(* IEC 61131-3 sources: SortJet_MasterSPS_Aufbau.fbsproj/08_POUs/Basis Funktionsbausteine, 5 files *)

(* ---- Ampel_FB.fb.st ---- *)
(* METADATA
{
	"v3Meta": {
		"objectGuid": "3b447e4d-6caa-4c98-ad2d-e4c3e81f2c59"
	}
}
*)
FUNCTION_BLOCK Ampel_FB
VAR_INPUT

  // BOOL
  bpAutomatikAktiv                : BOOL;
  bpSystemcheckAktiv              : BOOL;
  bpBetriebsstoppAktiv            : BOOL;
  bpInternerBetriebsstopp         : BOOL;
  bpHinweisFWEingriffErforderlich : BOOL;
  bpSignalExtern                  : BOOL; // Blau Dauerlicht (z. B. Faecherwagen bald voll); Eingriff erforderlich hat Vorrang (blinkt)

END_VAR
VAR_OUTPUT
END_VAR
VAR

  //BOOL
  blFlashbit    : BOOL;

  // BYTE
  bylShiftByte  : BYTE :=1;

  // WORD
  wlModus       : WORD;
  wlInitAmpel   : WORD;

  // INT
  ilIndex       : INT;

  // TRIGGER
  rtlInitAmpel  : R_TRIG;

  // BLINK
  Flasher       : BLINK;

END_VAR
VAR

  // HARDWARE AUSGAENGE
  out_bAmpelLeuchteRot     AT%Q* : BOOL;
  out_bAmpelLeuchteGelb    AT%Q* : BOOL;
  out_bAmpelLeuchteGruen   AT%Q* : BOOL;
  out_bAmpelLeuchteBlau    AT%Q* : BOOL;

END_VAR
//-------------------------------------------------------------------------------------------------
// BAUSTEIN: ANSTEUERUNG
//-------------------------------------------------------------------------------------------------
(* Hinweis:
   - Baustein zum Ansteuern der optischen Signale des Sortjet : AMPELN
*)
Flasher(ENABLE:= TRUE , TIMELOW:= t#0.2s, TIMEHIGH:= t#0.2s , OUT=> blFlashbit);
rtlInitAmpel(CLK:= blFlashbit );

out_bAmpelLeuchteBlau := SEL( bpHinweisFWEingriffErforderlich, bpSignalExtern, gbFlashbit02sec );

//  Zentral den OperatingMode bestimmen
IF ( NOT NotHalt.bpNotHaltOK) THEN // NotAus nicht OK
  wlModus := 3;
ELSIF ( bpBetriebsstoppAktiv  ) THEN // Betriebsstop gesetzt
  wlModus := 8;
ELSIF ( Visu_Start_Auto ) THEN // VisuAuto aktiv
  wlModus := 7;
ELSIF ( bgInbetriebnahmeBit ) THEN // Inbetriebnahmebit gesetzt
  wlModus := 5;
ELSIF ( bpInternerBetriebsstopp ) THEN // Fehler/interner betriebsstop gesetzt
  wlModus := 0;
ELSIF ( Initialisierung.bpInitialisierungAktiv ) THEN // Initialiesierung aktiv
  wlModus := 5;
ELSIF ( bpSystemcheckAktiv ) THEN // Checkroutine aktiv
  wlModus := 6;
ELSIF ( bpAutomatikAktiv ) THEN // automatik aktiv
  wlModus := 2;
ELSE // Handbetrieb aktiv
  wlModus := 4;
END_IF

CASE wlModus OF
  // ======================================================
  0 : // Faliure active
    out_bAmpelLeuchteRot    := blFlashbit;
    out_bAmpelLeuchteGelb   := NOT out_bAmpelLeuchteRot;
    out_bAmpelLeuchteGruen  := FALSE;

  // ======================================================
  1:  // Service Mode
    out_bAmpelLeuchteRot    := FALSE;
    out_bAmpelLeuchteGelb   := TRUE;
    out_bAmpelLeuchteGruen  := FALSE;

  // ======================================================
  2:  // Automatic Running
    out_bAmpelLeuchteRot    := FALSE;
    out_bAmpelLeuchteGelb   := FALSE;
    out_bAmpelLeuchteGruen  := TRUE;

  // ======================================================
  3:  // Emergency Stop Active
    out_bAmpelLeuchteRot    := TRUE;
    out_bAmpelLeuchteGelb   := FALSE;
    out_bAmpelLeuchteGruen  := FALSE;

  // ======================================================
  4:   // Manual Mode
    out_bAmpelLeuchteRot    := FALSE;
    out_bAmpelLeuchteGelb   := TRUE;
    out_bAmpelLeuchteGruen  := FALSE;

  // ======================================================
  5: // Initialisation Mode
    out_bAmpelLeuchteRot    := ((wlInitAmpel AND Maske_Bit_2)<>0);
    out_bAmpelLeuchteGelb   :=((wlInitAmpel AND Maske_Bit_1)<>0);
    out_bAmpelLeuchteGruen  :=((wlInitAmpel AND Maske_Bit_0)<>0);

  // ======================================================
  6:   // Check Routine wurde gestartet
    out_bAmpelLeuchteRot    := FALSE;
    out_bAmpelLeuchteGelb   := FALSE;
    out_bAmpelLeuchteGruen  := blFlashbit;

  // ======================================================
  7:   // VisuAuto aktiv
    out_bAmpelLeuchteRot    := FALSE;
    out_bAmpelLeuchteGelb   := NOT blFlashbit;
    out_bAmpelLeuchteGruen  := TRUE;
  // ======================================================
  8:   // Betriebsstoptaster betätigt
    out_bAmpelLeuchteRot    := FALSE;
    out_bAmpelLeuchteGelb   := blFlashbit;
    out_bAmpelLeuchteGruen  := bpAutomatikAktiv;

// ======================================================
END_CASE

IF ( wlModus = 5) THEN

  IF ( rtlInitAmpel.Q ) THEN

    wlInitAmpel :=SHL(bylShiftByte, ilIndex);
    ilIndex := ilIndex + 1;

    IF ( ilIndex = 3 ) THEN
      ilIndex := 0;
    END_IF;

  END_IF;

ELSE
  wlInitAmpel := 0;

END_IF
END_FUNCTION_BLOCK

(* ---- BetriebsStop_FB.fb.st ---- *)
(* METADATA
{
	"v3Meta": {
		"objectGuid": "07d57a24-f3c0-4742-8d44-44a8d21cf93a"
	}
}
*)
FUNCTION_BLOCK BetriebsStop_FB
VAR_INPUT
END_VAR
VAR_OUTPUT

  // BOOLEAN
  abpBetriebsstop  : ARRAY [cERSTER_AUTOMATIKKREIS..cLETZTER_AUTOMATIKKREIS] OF BOOL;

END_VAR
VAR

  // BOOLEAN
  blBetriebsstop  : BOOL; // Merkervariable

  // WORD
  wlIndex                    : WORD;
  wMeldungsNrInkrementieren  : WORD := 0;

END_VAR
//-------------------------------------------------------------------------------------------------
// BAUSTEIN: BETRIEBSSTATUS
//-------------------------------------------------------------------------------------------------

(* Hinweis:
   - Betriebs- Stopp ausloesen
   - Internen Betriebsstop ausloesen
*)

blBetriebsstop := (  ( NOT bgMMIOK AND NOT bgMMIBruecken ) );

//-------------------------------------------------------------------------------------------------
// BAUSTEIN: MELDUNGEN
//-------------------------------------------------------------------------------------------------
(* Hinweis:
   - Generieren einer Meldung
*)
wMeldungsNrInkrementieren := 0;

FOR wlIndex := cERSTER_AUTOMATIKKREIS TO cLETZTER_AUTOMATIKKREIS DO
  abpBetriebsstop[wlIndex] :=    Job_Stationen.abpFehler[wlIndex]
                                 OR Job_Shuttle.abpFehler[wlIndex]
                                 OR Job_Faecherwagen.abpFehler[wlIndex]
                                 OR NOT StatusAnlage.abpDruckluftOK[wlIndex]
                                 OR NOT StatusAnlage.bpAnlageOK
                                 OR blBetriebsstop;
  WatchIo( abpBetriebsstop[wlIndex] , ( ioccBetriebsstop1 + wMeldungsNrInkrementieren ) );
  wMeldungsNrInkrementieren := wMeldungsNrInkrementieren + 1;
END_FOR
END_FUNCTION_BLOCK

(* ---- Horn_FB.fb.st ---- *)
(* METADATA
{
	"v3Meta": {
		"objectGuid": "6f7ed93d-1901-4e95-8818-3caa484a7623"
	}
}
*)
FUNCTION_BLOCK Horn_FB
VAR_INPUT

  // BOOLEAN
  bpAktiv          : BOOL;
  bpReset          : BOOL;
  bpHornAktivieren : BOOL;  // Horn / Hupe vom Shuttle aus aktiviert

  // WORD
  wpStatusArt   : WORD; // Art des Hupsignales: 1=Dauerton 1; 2= Blinker 1/ 3= Blinker 2

  // TIME
  tpHornZeit   : TIME; // Zeit wie lange das Horn arbeitet

END_VAR
VAR_OUTPUT
END_VAR

VAR

  // BOOL
  blHornAktiv : BOOL;

  // TRIEGGER
  ftlHornAus  : F_TRIG;

  // TIMER
  tonlHornAus : TON;

END_VAR

VAR

  // HARDWAREAUSGAENGE
  out_bHorn       AT %Q* : BOOL; // akustische Anzeige, dass Checkroutine läuft

END_VAR

//-------------------------------------------------------------------------------------------------
// BAUSTEIN: ABLAUF HORNSIGNAL
//-------------------------------------------------------------------------------------------------
(* Hinweis:
   - Baustein zuruecksetzen
*)
IF ( bpReset  ) THEN

  bpReset    := FALSE;
  blHornAktiv := FALSE;

  out_bHorn  := FALSE;

ELSE

  (* Hinweis:
     - Aktivieren des Bausteins (Ablauf)
  *)
  IF ( bpAktiv ) THEN

    (* Hinweis:
       - Timer \ Trigger
    *)
    tonlHornAus(IN := blHornAktiv, PT:=tpHornZeit);

    ftlHornAus(CLK := blHornAktiv);

    IF ( bpHornAktivieren AND NOT blHornAktiv ) THEN
      blHornAktiv       := TRUE;
      bpHornAktivieren := FALSE;
    END_IF

    IF ( tonlHornAus.Q ) THEN
      blHornAktiv := FALSE;
    END_IF

    IF ( ftlHornAus.Q ) THEN
      out_bHorn := FALSE;
    END_IF

    (* Hinweis:
       - Hornsignal
    *)
    IF ( blHornAktiv ) THEN

      CASE wpStatusArt OF

        0,1:
          out_bHorn := TRUE;

        2:
          out_bHorn:= gbFlashbit1sec;

        3:
          out_bHorn:= gbFlashbit05sec;

        4:
          out_bHorn:= gbFlashbit02sec;

        5:
          out_bHorn:= gbFlashbit03sec;

        6:
          out_bHorn := gbFlashbit03sec AND gbFlashbit12sec;

        7:
          out_bHorn := gbFlashbit03sec AND gbFlashbit12sec;

      END_CASE

    ELSE
      out_bHorn  := FALSE;

    END_IF

  ELSE
    bpHornAktivieren := FALSE;
    out_bHorn := FALSE;

  END_IF

END_IF
END_FUNCTION_BLOCK

(* ---- PositionierAuftragsdatenPruefen.fb.st ---- *)
(* METADATA
{
	"v3Meta": {
		"objectGuid": "a4b12c85-33d1-4e58-8fdf-3218a4b905e2"
	}
}
*)
FUNCTION_BLOCK PositionierAuftragsdatenPruefen
VAR_INPUT

  rpSollPosition   : REAL; // Zielposition der Positionierung
  wpStationsNummer : WORD; // Station, die positioniert werden soll

END_VAR

VAR_OUTPUT

  // BOOLEAN
  bpErgebnis  : BOOL; // Rueckgabewert der Funktion

END_VAR

VAR

END_VAR
// Zentralestelle zum Ueberpruefen der Verfahrauftragsdaten [Positionieren]

bpErgebnis := TRUE;

Positionen();
END_FUNCTION_BLOCK

(* ---- Taktberechnung_FB.fb.st ---- *)
(* METADATA
{
	"v3Meta": {
		"objectGuid": "d72a9e43-2104-4490-bd51-13d6e7b9c79c"
	}
}
*)
FUNCTION_BLOCK Taktberechnung_FB
VAR_INPUT
  Signal             : BOOL;
END_VAR
VAR_OUTPUT
  Herz               : REAL;
END_VAR
VAR

  SignalSteigend     : R_TRIG;
  SignalFallend      : F_TRIG;

  tonZeitmessungOn   : TON;
  tonZeitmessungOff  : TON;

  tlOn               : TIME;
  tlOff              : TIME;
  tlHerz             : TIME;

END_VAR
SignalSteigend( CLK := Signal);
SignalFallend( CLK := Signal);

IF SignalSteigend.Q THEN
  tlOff := tonZeitmessungOff.ET;
END_IF

IF SignalFallend.Q THEN
  tlOn := tonZeitmessungOn.ET;
END_IF

tonZeitmessungOn( IN := Signal, PT := t#2s );
tonZeitmessungOff( IN := NOT Signal, PT := t#2s );

tlHerz := tlOff + tlOn;
IF tlHerz = T#0MS THEN
  tlHerz := T#1MS;
END_IF

IF NOT tonZeitmessungOff.Q AND NOT tonZeitmessungOn.Q THEN
  Herz := ( 1 / (TIME_TO_REAL(tlHerz) / 1000 ) );
ELSE
  Herz := 0.0;
END_IF
END_FUNCTION_BLOCK
